Fanuc KAREL source: KT00853.KL

PROGRAM KT00853
%NOLOCKGROUP
VAR
  B1: BOOLEAN
  B2: BOOLEAN
  OUT: REAL
BEGIN
  B1 = TRUE
  B2 = FALSE
  B1 = TRUE
  B2 = FALSE
  OUT = TAN(B1)
END KT00853
